(* IEC 61131-3 sources: sentinelot/zeek-lab/openplc-program, 1 file *)

(* ---- simple_plc.st ---- *)
PROGRAM plc_prg
  VAR
    counter_value AT %QW0 : INT;
  END_VAR

  counter_value := counter_value + 1;

END_PROGRAM

CONFIGURATION Config0

  RESOURCE Res0 ON PLC
    TASK task0(INTERVAL := T#20ms, PRIORITY := 0);
    PROGRAM instance0 WITH task0 : plc_prg;
  END_RESOURCE

END_CONFIGURATION
